    // NaN / 极大值保护，避免再次触发 FPU invalid。
    IF Yaw_W_enc_s <> Yaw_W_enc_s THEN
        Yaw_W_enc_s := 0.0;
        Yaw_W_last_enc_s := 0.0;
        Yaw_Alpha_enc_s2 := 0.0;
    ELSIF ABS(Yaw_W_enc_s) > Yaw_NumLimit_enc_s THEN
        Yaw_W_enc_s := 0.0;
        Yaw_W_last_enc_s := 0.0;
        Yaw_Alpha_enc_s2 := 0.0;
    END_IF;

    Yaw_Vraw_enc_s := Yaw_W_enc_s;
ELSE
    Yaw_W_enc_s := 0.0;
    Yaw_W_last_enc_s := 0.0;
    Yaw_Alpha_enc_s2 := 0.0;
    Yaw_Vraw_enc_s := 0.0;
END_IF;




// =============================================================
// T1. 机构学限位对力控 Vraw 的拦截
// 放在 U. 轴速度限幅之前；先判断，再进入速度/加速度/位置积分
// =============================================================
bLimitClampPlanar := FALSE;
bLimitClampAF := FALSE;

// BD 只受 CE-HI 限位
IF (BD_Vraw_enc_s > 0.0) AND bCEHI_Block_BD_Pos THEN
    BD_Vraw_enc_s := 0.0;
    bLimitClampPlanar := TRUE;
END_IF;

IF (BD_Vraw_enc_s < 0.0) AND bCEHI_Block_BD_Neg THEN
    BD_Vraw_enc_s := 0.0;
    bLimitClampPlanar := TRUE;
END_IF;

// AC 同时受 CAF 和 CE-HI 限位
IF (AC_Vraw_enc_s > 0.0) AND (bCAF_Block_AC_Pos OR bCEHI_Block_AC_Pos) THEN
    AC_Vraw_enc_s := 0.0;
    bLimitClampPlanar := TRUE;
END_IF;

IF (AC_Vraw_enc_s < 0.0) AND (bCAF_Block_AC_Neg OR bCEHI_Block_AC_Neg) THEN
    AC_Vraw_enc_s := 0.0;
    bLimitClampPlanar := TRUE;
END_IF;

// AF 同时受 CAF 和 CE-HI 限位
IF (AF_Vraw_enc_s > 0.0) AND (bCAF_Block_AF_Pos OR bCEHI_Block_AF_Pos) THEN
    AF_Vraw_enc_s := 0.0;
    bLimitClampAF := TRUE;
END_IF;

IF (AF_Vraw_enc_s < 0.0) AND (bCAF_Block_AF_Neg OR bCEHI_Block_AF_Neg) THEN
    AF_Vraw_enc_s := 0.0;
    bLimitClampAF := TRUE;
END_IF;

// 清导纳内部速度记忆，防止继续顶限位
IF bLimitClampPlanar THEN
    Vx_mps := 0.0;
    Vz_mps := 0.0;
    Vx_last_mps := 0.0;
    Vz_last_mps := 0.0;
    Ax_mps2 := 0.0;
    Az_mps2 := 0.0;
END_IF;

IF bLimitClampAF THEN
    AF_W_enc_s := 0.0;
    AF_W_last_enc_s := 0.0;
    AF_Alpha_enc_s2 := 0.0;
END_IF;


// =============================================================
// U. 轴速度限幅
// =============================================================
ScaleVel := 1.0;
ScaleVel_Axis := 1.0;

IF ABS(BD_Vraw_enc_s) > BD_Vmax_enc_s THEN
    tmpScale := BD_Vmax_enc_s / ABS(BD_Vraw_enc_s);
    IF tmpScale < ScaleVel THEN
        ScaleVel := tmpScale;
    END_IF;
END_IF;

IF ABS(AC_Vraw_enc_s) > AC_Vmax_enc_s THEN
    tmpScale := AC_Vmax_enc_s / ABS(AC_Vraw_enc_s);
    IF tmpScale < ScaleVel THEN
        ScaleVel := tmpScale;
    END_IF;
END_IF;

ScaleVel_Axis := ScaleVel;

BD_Vraw_enc_s := BD_Vraw_enc_s * ScaleVel_Axis;
AC_Vraw_enc_s := AC_Vraw_enc_s * ScaleVel_Axis;

// AF/Yaw 速度限幅：不用 x/ABS(x)，避免 Infinity/Infinity 触发 FPU invalid。
IF AF_Vraw_enc_s <> AF_Vraw_enc_s THEN
    AF_Vraw_enc_s := 0.0;
    AF_W_enc_s := 0.0;
    AF_W_last_enc_s := 0.0;
ELSIF ABS(AF_Vraw_enc_s) > AF_NumLimit_enc_s THEN
    AF_Vraw_enc_s := 0.0;
    AF_W_enc_s := 0.0;
    AF_W_last_enc_s := 0.0;
END_IF;

IF AF_Vraw_enc_s > AF_Vmax_enc_s THEN
    AF_Vraw_enc_s := AF_Vmax_enc_s;
ELSIF AF_Vraw_enc_s < -AF_Vmax_enc_s THEN
    AF_Vraw_enc_s := -AF_Vmax_enc_s;
END_IF;

IF Yaw_Vraw_enc_s <> Yaw_Vraw_enc_s THEN
    Yaw_Vraw_enc_s := 0.0;
    Yaw_W_enc_s := 0.0;
    Yaw_W_last_enc_s := 0.0;
ELSIF ABS(Yaw_Vraw_enc_s) > 100000.0 THEN
    Yaw_Vraw_enc_s := 0.0;
    Yaw_W_enc_s := 0.0;
    Yaw_W_last_enc_s := 0.0;
END_IF;

IF Yaw_Vraw_enc_s > Yaw_Vmax_enc_s THEN
    Yaw_Vraw_enc_s := Yaw_Vmax_enc_s;
ELSIF Yaw_Vraw_enc_s < -Yaw_Vmax_enc_s THEN
    Yaw_Vraw_enc_s := -Yaw_Vmax_enc_s;
END_IF;


// =============================================================
// V. 加速度限幅
// =============================================================
BD_Vlast_enc_s := BD_Vcmd_enc_s;
AC_Vlast_enc_s := AC_Vcmd_enc_s;
AF_Vlast_enc_s := AF_Vcmd_enc_s;
Yaw_Vlast_enc_s := Yaw_Vcmd_enc_s;

// AC/BD 加减速度限幅：
// 1) 加速使用 BD_Amax/AC_Amax；
// 2) 撤力减速或反向使用 BD_Dmax/AC_Dmax；
// 3) 最后用同一个 ScaleAcc_Axis 同步缩放 BD/AC，保持末端方向不被破坏。
BD_dV_enc_s := BD_Vraw_enc_s - BD_Vlast_enc_s;
AC_dV_enc_s := AC_Vraw_enc_s - AC_Vlast_enc_s;

IF (ABS(BD_Vraw_enc_s) < ABS(BD_Vlast_enc_s)) OR (BD_Vraw_enc_s * BD_Vlast_enc_s < 0.0) THEN
    BD_dVmax_enc_s := BD_Dmax_enc_s2 * Ts;
ELSE
    BD_dVmax_enc_s := BD_Amax_enc_s2 * Ts;
END_IF;

IF (ABS(AC_Vraw_enc_s) < ABS(AC_Vlast_enc_s)) OR (AC_Vraw_enc_s * AC_Vlast_enc_s < 0.0) THEN
    AC_dVmax_enc_s := AC_Dmax_enc_s2 * Ts;
ELSE
    AC_dVmax_enc_s := AC_Amax_enc_s2 * Ts;
END_IF;

ScaleAcc := 1.0;
ScaleAcc_Axis := 1.0;

IF ABS(BD_dV_enc_s) > BD_dVmax_enc_s THEN
    IF BD_dVmax_enc_s > 0.0 THEN
        tmpScale := BD_dVmax_enc_s / ABS(BD_dV_enc_s);
    ELSE
        tmpScale := 0.0;
    END_IF;
    IF tmpScale < ScaleAcc THEN
        ScaleAcc := tmpScale;
    END_IF;
END_IF;

IF ABS(AC_dV_enc_s) > AC_dVmax_enc_s THEN
    IF AC_dVmax_enc_s > 0.0 THEN
        tmpScale := AC_dVmax_enc_s / ABS(AC_dV_enc_s);
    ELSE
        tmpScale := 0.0;
    END_IF;
    IF tmpScale < ScaleAcc THEN
        ScaleAcc := tmpScale;
    END_IF;
END_IF;

ScaleAcc_Axis := ScaleAcc;

BD_Vcmd_enc_s := BD_Vlast_enc_s + BD_dV_enc_s * ScaleAcc_Axis;
AC_Vcmd_enc_s := AC_Vlast_enc_s + AC_dV_enc_s * ScaleAcc_Axis;

IF Ts > 0.000001 THEN
    BD_Acmd_enc_s2 := (BD_Vcmd_enc_s - BD_Vlast_enc_s) / Ts;
    AC_Acmd_enc_s2 := (AC_Vcmd_enc_s - AC_Vlast_enc_s) / Ts;
ELSE
    BD_Acmd_enc_s2 := 0.0;
    AC_Acmd_enc_s2 := 0.0;
END_IF;

// AF 加减速度限幅：加速用 AF_Amax，撤力减速/反向用更大的 AF_Dmax。
AF_dV_enc_s := AF_Vraw_enc_s - AF_Vlast_enc_s;

IF (ABS(AF_Vraw_enc_s) < ABS(AF_Vlast_enc_s)) OR (AF_Vraw_enc_s * AF_Vlast_enc_s < 0.0) THEN
    AF_dVmax_enc_s := AF_Dmax_enc_s2 * Ts;
ELSE
    AF_dVmax_enc_s := AF_Amax_enc_s2 * Ts;
END_IF;

IF AF_dV_enc_s > AF_dVmax_enc_s THEN
    AF_dV_enc_s := AF_dVmax_enc_s;
ELSIF AF_dV_enc_s < -AF_dVmax_enc_s THEN
    AF_dV_enc_s := -AF_dVmax_enc_s;
END_IF;

AF_Vcmd_enc_s := AF_Vlast_enc_s + AF_dV_enc_s;

IF Ts > 0.000001 THEN
    AF_Acmd_enc_s2 := (AF_Vcmd_enc_s - AF_Vlast_enc_s) / Ts;
ELSE
    AF_Acmd_enc_s2 := 0.0;
END_IF;

// yaw 加减速度限幅：加速用 Yaw_Amax，撤力减速/反向用 Yaw_Dmax。
Yaw_dV_enc_s := Yaw_Vraw_enc_s - Yaw_Vlast_enc_s;

IF (ABS(Yaw_Vraw_enc_s) < ABS(Yaw_Vlast_enc_s)) OR (Yaw_Vraw_enc_s * Yaw_Vlast_enc_s < 0.0) THEN
    Yaw_dVmax_enc_s := Yaw_Dmax_enc_s2 * Ts;
ELSE
    Yaw_dVmax_enc_s := Yaw_Amax_enc_s2 * Ts;
END_IF;

IF Yaw_dV_enc_s > Yaw_dVmax_enc_s THEN
    Yaw_dV_enc_s := Yaw_dVmax_enc_s;
ELSIF Yaw_dV_enc_s < -Yaw_dVmax_enc_s THEN
    Yaw_dV_enc_s := -Yaw_dVmax_enc_s;
END_IF;

Yaw_Vcmd_enc_s := Yaw_Vlast_enc_s + Yaw_dV_enc_s;

IF Ts > 0.000001 THEN
    Yaw_Acmd_enc_s2 := (Yaw_Vcmd_enc_s - Yaw_Vlast_enc_s) / Ts;
ELSE
    Yaw_Acmd_enc_s2 := 0.0;
END_IF;




// =============================================================
// V1. 机构学限位对力控 Vcmd 的最终保险
// 放在 W. 小速度归零之前，位置积分之前
// =============================================================
// BD
IF (BD_Vcmd_enc_s > 0.0) AND bCEHI_Block_BD_Pos THEN
    BD_Vcmd_enc_s := 0.0;
    BD_Acmd_enc_s2 := 0.0;
END_IF;

IF (BD_Vcmd_enc_s < 0.0) AND bCEHI_Block_BD_Neg THEN
    BD_Vcmd_enc_s := 0.0;
    BD_Acmd_enc_s2 := 0.0;
END_IF;

// AC
IF (AC_Vcmd_enc_s > 0.0) AND (bCAF_Block_AC_Pos OR bCEHI_Block_AC_Pos) THEN
    AC_Vcmd_enc_s := 0.0;
    AC_Acmd_enc_s2 := 0.0;
END_IF;

IF (AC_Vcmd_enc_s < 0.0) AND (bCAF_Block_AC_Neg OR bCEHI_Block_AC_Neg) THEN
    AC_Vcmd_enc_s := 0.0;
    AC_Acmd_enc_s2 := 0.0;
END_IF;

// AF
IF (AF_Vcmd_enc_s > 0.0) AND (bCAF_Block_AF_Pos OR bCEHI_Block_AF_Pos) THEN
    AF_Vcmd_enc_s := 0.0;
    AF_Acmd_enc_s2 := 0.0;
    AF_W_enc_s := 0.0;
    AF_W_last_enc_s := 0.0;
END_IF;

IF (AF_Vcmd_enc_s < 0.0) AND (bCAF_Block_AF_Neg OR bCEHI_Block_AF_Neg) THEN
    AF_Vcmd_enc_s := 0.0;
    AF_Acmd_enc_s2 := 0.0;
    AF_W_enc_s := 0.0;
    AF_W_last_enc_s := 0.0;
END_IF;


// =============================================================
// W. 小速度归零
// =============================================================
IF ABS(BD_Vcmd_enc_s) < 0.001 THEN
    BD_Vcmd_enc_s := 0.0;
END_IF;

IF ABS(AC_Vcmd_enc_s) < 0.001 THEN
    AC_Vcmd_enc_s := 0.0;
END_IF;

IF ABS(AF_Vcmd_enc_s) < 0.02 THEN
    AF_Vcmd_enc_s := 0.0;
END_IF;

IF ABS(Yaw_Vcmd_enc_s) < 0.001 THEN
    Yaw_Vcmd_enc_s := 0.0;
END_IF;

// =============================================================
// W1. 轴1抱闸未释放时冻结 BD 给定
// 防止抱闸合上或释放延时未到时，BD 外部位置继续积分。
// =============================================================
IF NOT Axis1_BrakeMotionOK THEN
    BD_Vraw_enc_s := 0.0;
    BD_Vcmd_enc_s := 0.0;
    BD_Vlast_enc_s := 0.0;
    BD_Acmd_enc_s2 := 0.0;
    qdotBD_m_s := 0.0;
    BD_PosCmd_Enc := BD_ActEnc;
END_IF;


// =============================================================
// X. 力控基础软限位
// 当前只对 axis1=BD 编码器 2~600 做限位
// =============================================================
bForceSoftLimit := FALSE;

BD_NextCmd_Enc := BD_PosCmd_Enc + BD_Vcmd_enc_s * Ts;
AC_NextCmd_Enc := AC_PosCmd_Enc + AC_Vcmd_enc_s * Ts;
AF_NextCmd_Enc := AF_PosCmd_Enc + AF_Vcmd_enc_s * Ts;
Yaw_NextCmd_Enc := Yaw_PosCmd_Enc + Yaw_Vcmd_enc_s * Ts;

IF (BD_NextCmd_Enc < BD_EncMin) OR (BD_NextCmd_Enc > BD_EncMax) THEN
    bForceSoftLimit := TRUE;
END_IF;

IF bUseAFLimit THEN
    IF (AF_NextCmd_Enc < AF_EncMin) OR (AF_NextCmd_Enc > AF_EncMax) THEN
        bForceSoftLimit := TRUE;
    END_IF;
END_IF;

IF (Yaw_NextCmd_Enc < Base_EncMin) OR (Yaw_NextCmd_Enc > Base_EncMax) THEN
    bForceSoftLimit := TRUE;
END_IF;

IF bForceSoftLimit THEN
    BD_Vcmd_enc_s := 0.0;
    AC_Vcmd_enc_s := 0.0;
    AF_Vcmd_enc_s := 0.0;
    Yaw_Vcmd_enc_s := 0.0;

    BD_Acmd_enc_s2 := 0.0;
    AC_Acmd_enc_s2 := 0.0;
    AF_Acmd_enc_s2 := 0.0;
    Yaw_Acmd_enc_s2 := 0.0;

    Vx_mps := 0.0;
    Vz_mps := 0.0;
    AF_W_enc_s := 0.0;
    Yaw_W_enc_s := 0.0;
END_IF;


// =============================================================
// Y. 位置积分
// 外部位置给定使用真实 NC 编码器坐标
// =============================================================
IF bRunForce AND NOT bForceSoftLimit THEN
    BD_PosCmd_Enc := BD_PosCmd_Enc + BD_Vcmd_enc_s * Ts;
    AC_PosCmd_Enc := AC_PosCmd_Enc + AC_Vcmd_enc_s * Ts;
    AF_PosCmd_Enc := AF_PosCmd_Enc + AF_Vcmd_enc_s * Ts;
    Yaw_PosCmd_Enc := Yaw_PosCmd_Enc + Yaw_Vcmd_enc_s * Ts;
END_IF;


// =============================================================
// Z. Direction 判断
// =============================================================
IF BD_Vcmd_enc_s > 0.001 THEN
    DirBD := 1;
ELSIF BD_Vcmd_enc_s < -0.001 THEN
    DirBD := -1;
ELSE
    DirBD := 0;
END_IF;

IF AC_Vcmd_enc_s > 0.001 THEN
    DirAC := 1;
ELSIF AC_Vcmd_enc_s < -0.001 THEN
    DirAC := -1;
ELSE
    DirAC := 0;
END_IF;

IF AF_Vcmd_enc_s > 0.001 THEN
    DirAF := 1;
ELSIF AF_Vcmd_enc_s < -0.001 THEN
    DirAF := -1;
ELSE
    DirAF := 0;
END_IF;

IF Yaw_Vcmd_enc_s > 0.001 THEN
    DirYaw := 1;
ELSIF Yaw_Vcmd_enc_s < -0.001 THEN
    DirYaw := -1;
ELSE
    DirYaw := 0;
END_IF;


// =============================================================
// Z1. 每周期 Feed axis1 / axis2 / axis3 / axis4
// 急停、未 Ready、未力控时，不再 Feed，避免恢复后继续追旧目标。
// =============================================================
IF bRunForce AND bAxesReadyForForce THEN
    bFeedBD := MC_ExtSetPointGenFeed(
        Axis := axis1,
        Position := BD_PosCmd_Enc,
        Velocity := ABS(BD_Vcmd_enc_s),
        Acceleration := ABS(BD_Acmd_enc_s2),
        Direction := DirBD
    );

    bFeedAC := MC_ExtSetPointGenFeed(
        Axis := axis2,
        Position := AC_PosCmd_Enc,
        Velocity := ABS(AC_Vcmd_enc_s),
        Acceleration := ABS(AC_Acmd_enc_s2),
        Direction := DirAC
    );

    bFeedAF := MC_ExtSetPointGenFeed(
        Axis := axis3,
        Position := AF_PosCmd_Enc,
        Velocity := ABS(AF_Vcmd_enc_s),
        Acceleration := ABS(AF_Acmd_enc_s2),
        Direction := DirAF
    );

    bFeedYaw := MC_ExtSetPointGenFeed(
        Axis := axis4,
        Position := Yaw_PosCmd_Enc,
        Velocity := ABS(Yaw_Vcmd_enc_s),
        Acceleration := ABS(Yaw_Acmd_enc_s2),
        Direction := DirYaw
    );
ELSE
    bFeedBD := FALSE;
    bFeedAC := FALSE;
    bFeedAF := FALSE;
    bFeedYaw := FALSE;

    // 非力控/急停/轴未 Ready 时保持目标等于当前位置，防止恢复后跳变。
    IF NOT bRunForce THEN
        BD_PosCmd_Enc := BD_ActEnc;
        AC_PosCmd_Enc := AC_ActEnc;
        AF_PosCmd_Enc := AF_ActEnc;
        Yaw_PosCmd_Enc := Yaw_ActEnc;
    END_IF;
END_IF;


// =============================================================
// Z2. 抱闸和灯
// =============================================================
// 轴1抱闸 axis1baozha 已在 D1 中按“轴1真实使能 + 无故障 + 300ms 延时”逻辑处理。
// 这里保留 axis4 原逻辑。注意：axis4 不受 CE-HI 限位影响。
axis4baozha := ballow_axis4jogfw OR ballow_axis4jogbw OR bRunForce;

// 电磁阀和电磁阀灯完全独立，不经过 CAF/CEHI 限位。
valveopen1 := valvejudge;
valveopen2 := valvejudge;
valvelight := valvejudge;

// 指示灯也从 CEHI/CAF 限位逻辑中拆出来：
// 手动模式下，只要按钮输入为 TRUE 就亮，用于确认按钮链路；
// 力控模式下，对应轴有速度给定时也亮。
// 这样即使某方向被软限位禁止，按键灯仍能亮，便于判断“输入有效但被限位拦截”。
bOutput_axis1light :=
    bInput_axis1jogfw OR bInput_axis1jogbw
    OR (bRunForce AND (ABS(BD_Vcmd_enc_s) > 0.001));

bOutput_axis2light :=
    bInput_axis2jogfw OR bInput_axis2jogbw
    OR (bRunForce AND (ABS(AC_Vcmd_enc_s) > 0.001));

bOutput_axis3light :=
    bInput_axis3jogfw OR bInput_axis3jogbw
    OR (bRunForce AND (ABS(AF_Vcmd_enc_s) > 0.02));

bOutput_axis4light :=
    bInput_axis4jogfw OR bInput_axis4jogbw
    OR (bRunForce AND (ABS(Yaw_Vcmd_enc_s) > 0.001));

    likonglight := bForceMode;

// =============================================================
// Z3. 错误输出
// =============================================================
axis1_status(Axis := axis1, Enable := TRUE);
axis2_status(Axis := axis2, Enable := TRUE);
axis3_status(Axis := axis3, Enable := TRUE);
axis4_status(Axis := axis4, Enable := TRUE);

bAxis1Err := axis1_power.Error OR axis1_status.Error OR axis1_status.ErrorStop;
bAxis2Err := axis2_power.Error OR axis2_status.Error OR axis2_status.ErrorStop;
bAxis3Err := axis3_power.Error OR axis3_status.Error OR axis3_status.ErrorStop;
bAxis4Err := axis4_power.Error OR axis4_status.Error OR axis4_status.ErrorStop;

bAnyAxisErr := bAxis1Err OR bAxis2Err OR bAxis3Err OR bAxis4Err;

IF bResetStopReason THEN
    StopReasonCode := 0;
    bStopReasonLatched := FALSE;
END_IF;

IF bRunForce AND NOT bStopReasonLatched THEN

    IF NOT bForceMode THEN
        StopReasonCode := 1;
        bStopReasonLatched := TRUE;

    ELSIF NOT bAxesReadyForForce THEN
        StopReasonCode := 2;
        bStopReasonLatched := TRUE;

   ELSIF bAnyAxisErr THEN
    StopReasonCode := 3;
    bStopReasonLatched := TRUE;
    

    ELSIF bCEHI_Block_BD_Pos OR bCEHI_Block_BD_Neg
       OR bCEHI_Block_AC_Pos OR bCEHI_Block_AC_Neg
       OR bCEHI_Block_AF_Pos OR bCEHI_Block_AF_Neg THEN
        StopReasonCode := 4;
        bStopReasonLatched := TRUE;

    ELSIF bCAF_Block_AC_Pos OR bCAF_Block_AC_Neg
       OR bCAF_Block_AF_Pos OR bCAF_Block_AF_Neg THEN
        StopReasonCode := 5;
        bStopReasonLatched := TRUE;

    ELSIF NOT bExtBD OR NOT bExtAC THEN
        StopReasonCode := 6;
        bStopReasonLatched := TRUE;

    ELSIF NOT Axis1_BrakeMotionOK THEN
        StopReasonCode := 7;
        bStopReasonLatched := TRUE;
    END_IF;

END_IF;

bError := axis1_power.Error OR axis2_power.Error OR axis3_power.Error OR axis4_power.Error
       OR axis1_jogerror OR axis2_jogerror OR axis3_jogerror OR axis4_jogerror
       OR fbExtEnableBD.Error OR fbExtEnableAC.Error OR fbExtEnableAF.Error OR fbExtEnableYaw.Error
       OR fbExtDisableBD.Error OR fbExtDisableAC.Error OR fbExtDisableAF.Error OR fbExtDisableYaw.Error
       OR axis1_reset.Error OR axis2_reset.Error OR axis3_reset.Error OR axis4_reset.Error;

IF axis1_power.Error THEN
    nErrorID := axis1_power.ErrorID;
ELSIF axis2_power.Error THEN
    nErrorID := axis2_power.ErrorID;
ELSIF axis3_power.Error THEN
    nErrorID := axis3_power.ErrorID;
ELSIF axis4_power.Error THEN
    nErrorID := axis4_power.ErrorID;
ELSIF axis1_jogerror THEN
    nErrorID := axis1_jogerrorid;
ELSIF axis2_jogerror THEN
    nErrorID := axis2_jogerrorid;
ELSIF axis3_jogerror THEN
    nErrorID := axis3_jogerrorid;
ELSIF axis4_jogerror THEN
    nErrorID := axis4_jogerrorid;
ELSIF fbExtEnableBD.Error THEN
    nErrorID := fbExtEnableBD.ErrorID;
ELSIF fbExtEnableAC.Error THEN
    nErrorID := fbExtEnableAC.ErrorID;
ELSIF fbExtEnableAF.Error THEN
    nErrorID := fbExtEnableAF.ErrorID;
ELSIF fbExtEnableYaw.Error THEN
    nErrorID := fbExtEnableYaw.ErrorID;
ELSIF fbExtDisableBD.Error THEN
    nErrorID := fbExtDisableBD.ErrorID;
ELSIF fbExtDisableAC.Error THEN
    nErrorID := fbExtDisableAC.ErrorID;
ELSIF fbExtDisableAF.Error THEN
    nErrorID := fbExtDisableAF.ErrorID;
ELSIF fbExtDisableYaw.Error THEN
    nErrorID := fbExtDisableYaw.ErrorID;
ELSIF axis1_reset.Error THEN
    nErrorID := axis1_reset.ErrorID;
ELSIF axis2_reset.Error THEN
    nErrorID := axis2_reset.ErrorID;
ELSIF axis3_reset.Error THEN
    nErrorID := axis3_reset.ErrorID;
ELSIF axis4_reset.Error THEN
    nErrorID := axis4_reset.ErrorID;
ELSE
    nErrorID := 0;
END_IF;

END_PROGRAM

(* stored: Version 1.1.0.1, ProductVersion 3.1.4024.16
   POU MAIN: Id {81832343-112e-4f9b-82f5-774ce7357d5e}, SpecialFunc None *)
